TYPE ST_MUNSCH_REF : FB_MUNSCH_EXTRUDER_REF;
END_TYPE

(* stored: Version 1.1.0.1, ProductVersion 3.1.4024.15
   DUT ST_MUNSCH_REF: Id {232061af-a530-4698-9a44-1a2f3f5cecc8} *)
